// TIA Portal V21 export
// export: Created 2026-11-10T20:11:28.2910772Z, ExportSetting WithDefaults, DisplayName Totally Integrated Automation Portal, DisplayVersion V21 Update 3, DisplayName STEP 7 Professional, DisplayVersion V21 Update 3, DisplayName STEP 7 Safety, DisplayVersion V21, DisplayName Tech WebApplication, DisplayVersion V21, DisplayName WinCC Basic/Comfort/Advanced, DisplayVersion V21 Update 3, DisplayName WinCC Unified, DisplayVersion V21 Update 3
FUNCTION_BLOCK "FB_FbdStruct"   // FB100, FBD
{ S7_Optimized_Access := 'TRUE' }
VERSION : 0.1
// stored: AutoNumber true, IsIECCheckEnabled false, IsRetainMemResEnabled false, MemoryReserve 100, SetENOAutomatically false, UDAEnableTagReadback false
   VAR_INPUT
      "a" : Bool;
      "b" : Bool;
      c : Bool;
      ia : Int;
   END_VAR
   VAR_OUTPUT
      q : Bool;
      q2 : Bool;
      io : Int;
      io2 : Int;
   END_VAR
   VAR
      ifc1 { S7_SetPoint := 'True'} : "FB_Iface";
      ton1 { S7_SetPoint := 'True'} : TON_TIME;
   END_VAR
BEGIN

REGION Network 1: AND then OR
   // Gate cascade
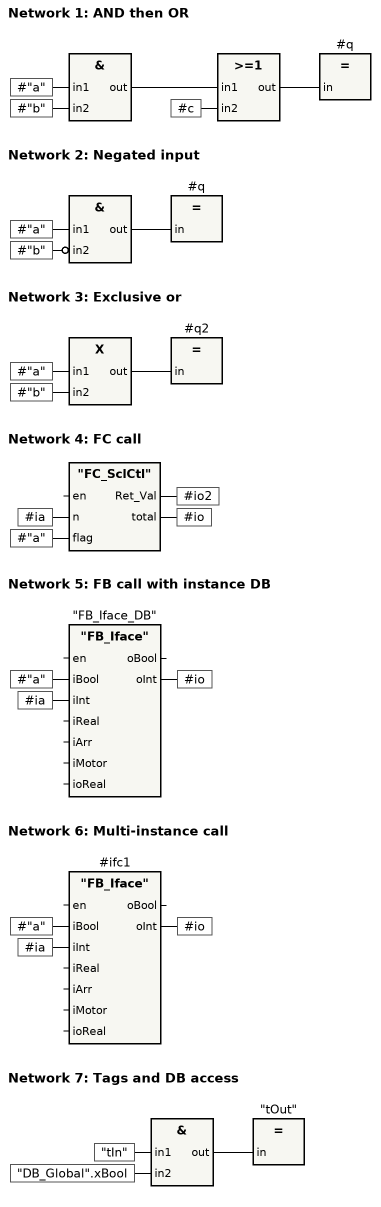
   #q := (#"a" AND #"b") OR #c;
END_REGION

REGION Network 2: Negated input
   #q := #"a" AND NOT #"b";
END_REGION

REGION Network 3: Exclusive or
   #q2 := #"a" XOR #"b";
END_REGION

REGION Network 4: FC call
   #io2 := "FC_SclCtl"(n := #ia, flag := #"a", total => #io);
END_REGION

REGION Network 5: FB call with instance DB
   "FB_Iface_DB"(iBool := #"a", iInt := #ia, oInt => #io);   // "FB_Iface"
END_REGION

REGION Network 6: Multi-instance call
   #ifc1(iBool := #"a", iInt := #ia, oInt => #io);   // "FB_Iface"
END_REGION

REGION Network 7: Tags and DB access
   "tOut" := "tIn" AND "DB_Global".xBool;
END_REGION
END_FUNCTION_BLOCK
